TYPE ET_ItpWriteRParams :
(
	ET_ItpWriteRParams_eWaitExecute := 0,
	ET_ItpWriteRParams_eWriteRParams := 5,
	ET_ItpWriteRParams_eDone := 197,
	ET_ItpWriteRParams_eError := 198,
	ET_ItpWriteRParams_eNoExecute := 199
);
END_TYPE

(* stored: Version 1.1.0.1, ProductVersion 3.1.4024.15
   DUT ET_ItpWriteRParams: Id {231e1fad-5b9d-4e22-a02f-e0e4d1857235} *)
